FUNCTION_BLOCK ESP32_OPCUA_SERVER_1 (* Starts the ESP32 OPC UA server *)
  (* Standard: 61499-2; Description: ESP32 OPC UA server control block *)
  (* Version 1.0, 2026-11-23, Jose Helio, Esp Forte OPC UA, Server control service interface function block *)
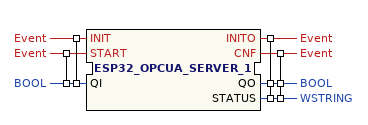
  EVENT_INPUT
    INIT WITH QI; (* Initialize the block *)
    START WITH QI; (* Start the OPC UA server *)
  END_EVENT
  EVENT_OUTPUT
    INITO WITH QO, STATUS; (* Initialization confirmation *)
    CNF WITH QO, STATUS; (* Start confirmation *)
  END_EVENT
  VAR_INPUT
    QI : BOOL; (* Enable the service *)
  END_VAR
  VAR_OUTPUT
    QO : BOOL; (* Operation result *)
    STATUS : WSTRING; (* Server status *)
  END_VAR
END_FUNCTION_BLOCK
